(* IEC 61131-3 sources: 2026_Projet_YGO_ExcavatriceDragage/ARCHIVES/Code/MAIN, 3 files *)

(* ---- PRG_01_Inputs_LD.st ---- *)
(* ═══════════════════════════════════════════════════════════════
   📥 PRG_01_Inputs_LD — ACQUISITION & QUALIFICATION DES ENTRÉES (LADDER)
   ───────────────────────────────────────────────────────────────
   📄 Doc : DOC/AF_Partie-06_Acquisition_Qualification_IO_v2.1.md §1/§4
   ⚙️ Exécuté par la tâche PLC en position 1 (premier programme).
   🎯 Lit les 22 TOR réelles depuis leurs symboles bruts mappés (CSV
       Device_IO_20260729.csv), applique un filtre anti-rebond 20 ms et
       publie :
         • Qualified : ST_InputsQualified  (image qualifiée, lecteur unique
                                            PRG_02_Acquisition_CFC)
         • 14 scalaires legacy             (consommateurs historiques)
   🛡️ Polarité : le nom de chaque entrée dit ce que TRUE signifie. Seuls
       les freins portent InvertLogic := FALSE (REX 2026-08-03 : TRUE =
       frein OUVERT). Aucune autre inversion (contacts NC câblés 1 = sain).
   📄 Converti automatiquement en Ladder Diagram (<LD>) dans CODESYS.
   ═══════════════════════════════════════════════════════════════ *)

PROGRAM PRG_01_Inputs_LD
VAR_OUTPUT
    Qualified : ST_InputsQualified;
    PowerContactorEngaged : BOOL;   // TRUE = contacteur de puissance engagé (NO)
    EmergencyChainClosed  : BOOL;   // TRUE = boucle AU fermée (NC, câblage 1 = sain)
    PhaseRotationOk       : BOOL;   // TRUE = rotation phases correcte (NC)
    BrakeThermalFeedback  : BOOL;   // TRUE = thermique freins M1/M2/M3 OK (NC)
    M1ThermalFeedback     : BOOL;   // TRUE = thermique M1 OK (NC)
    M2ThermalFeedback     : BOOL;   // TRUE = thermique M2 OK (NC)
    M1BrakeFeedback       : BOOL;   // TRUE = frein M1 OUVERT (desserré) — REX 2026-08-03
    M2BrakeFeedback       : BOOL;   // TRUE = frein M2 OUVERT (desserré) — REX 2026-08-03
    M3BrakeFeedback       : BOOL;   // TRUE = frein M3 OUVERT (desserré) — REX 2026-08-03
    M1FwdRevSpeedFeedbackOff : BOOL; // TRUE = contacteurs sens M1 retombés (NO)
    M2FwdRevSpeedFeedbackOff : BOOL; // TRUE = contacteurs sens M2 retombés (NO)
    TopPositionSensor     : BOOL;   // TRUE = position extrême haut libre (NC)
    SlackCableSwitch      : BOOL;   // TRUE = câble M2 tendu (NC)
    KoboldContactFond     : BOOL;   // TRUE = Kobold fond détecté (NO)
END_VAR
VAR
    instPowerContactorEngaged : FB_Input;
    instEmergencyChainClosed  : FB_Input;
    instCtrlPhaseRotation     : FB_Input;
    instBrakeThermalFeedback  : FB_Input;
    instKoboldContactFond     : FB_Input;
    instHydraulicThermalOk    : FB_Input;
    instConveyorInfeedReady   : FB_Input;
    instM1FwdRevSpeedFeedbackOff : FB_Input;
    instM1Thermal             : FB_Input;
    instM1BrakeFeedback       : FB_Input;
    instM2FwdRevSpeedFeedbackOff : FB_Input;
    instM2Thermal             : FB_Input;
    instM2BrakeFeedback       : FB_Input;
    instTopPositionSensor     : FB_Input;
    instSlackCableSwitch      : FB_Input;
    instM3BrakeFeedback       : FB_Input;
    instM3ThermalFeedback     : FB_Input;
    instTranslationPosTremie  : FB_Input;
    instTranslationPosPV      : FB_Input;
    instTranslationPosP2      : FB_Input;
    instTranslationPosP1      : FB_Input;
    instTranslationPosMaintenance : FB_Input;
END_VAR

// === IMPLEMENTATION ===

// === [MACHINE] ===
// 🔌 Contacteur de puissance géré par l'arrêt d'urgence (NO) — TRUE = engagé
instPowerContactorEngaged(InputRaw := PowerContactorEngaged_DI, FilterTime := T#20MS);
PowerContactorEngaged := instPowerContactorEngaged.State;
Qualified.Machine.PowerContactorEngaged_DI := PowerContactorEngaged;

// 🔗 Boucle d'arrêt d'urgence coup-de-poing + contact PLC (NC) — TRUE = saine
instEmergencyChainClosed(InputRaw := EmergencyChainClosed_DI, FilterTime := T#20MS);
EmergencyChainClosed := instEmergencyChainClosed.State;
Qualified.Machine.EmergencyChainClosed_DI := EmergencyChainClosed;

// ⚡ Contrôle rotation phases (NC) — TRUE = correcte
instCtrlPhaseRotation(InputRaw := PhaseRotationOk_DI, FilterTime := T#20MS);
PhaseRotationOk := instCtrlPhaseRotation.State;
Qualified.Machine.PhaseRotationOk_DI := PhaseRotationOk;

// 🌡️ Thermique freins commun M1/M2/M3 (NC) — TRUE = OK
instBrakeThermalFeedback(InputRaw := BrakeThermalOk_DI, FilterTime := T#20MS);
BrakeThermalFeedback := instBrakeThermalFeedback.State;
Qualified.Machine.BrakeThermalOk_DI := BrakeThermalFeedback;

// 🪨 Détecteur fond Kobold (NO) — TRUE = fond détecté
instKoboldContactFond(InputRaw := M1_M2_KoboldContactFond_DI, FilterTime := T#20MS);
KoboldContactFond := instKoboldContactFond.State;
Qualified.Machine.M1_M2_KoboldContactFond_DI := KoboldContactFond;

// 🌡️ Thermique moteur hydraulique (NC) — TRUE = OK
instHydraulicThermalOk(InputRaw := HydraulicThermalOk_DI, FilterTime := T#20MS);
Qualified.Machine.HydraulicThermalOk_DI := instHydraulicThermalOk.State;

// ⚙️ Autorisation démarrage crible (NO) — TRUE = autorisé
instConveyorInfeedReady(InputRaw := ConveyorInfeedReady_DI, FilterTime := T#20MS);
Qualified.Machine.ConveyorInfeedReady_DI := instConveyorInfeedReady.State;

// === [WINCH] ===
// 📡 Contacteurs sens M1 relâchés (NO) — TRUE = retombés
instM1FwdRevSpeedFeedbackOff(InputRaw := M1_ContactorsReleased_DI, FilterTime := T#20MS);
M1FwdRevSpeedFeedbackOff := instM1FwdRevSpeedFeedbackOff.State;
Qualified.Winch.M1_ContactorsReleased_DI := M1FwdRevSpeedFeedbackOff;

// 🌡️ Thermique moteur M1 (NC) — TRUE = OK
instM1Thermal(InputRaw := M1_ThermalOk_DI, FilterTime := T#20MS);
M1ThermalFeedback := instM1Thermal.State;
Qualified.Winch.M1_ThermalOk_DI := M1ThermalFeedback;

// 🔒 Retour frein M1 — REX 2026-08-03 : InvertLogic := FALSE, TRUE = frein OUVERT
instM1BrakeFeedback(InputRaw := M1_BrakeIsOpen_DI, InvertLogic := FALSE, FilterTime := T#20MS);
M1BrakeFeedback := instM1BrakeFeedback.State;
Qualified.Winch.M1_BrakeIsOpen_DI := M1BrakeFeedback;

// 📡 Contacteurs sens M2 relâchés (NO) — TRUE = retombés
instM2FwdRevSpeedFeedbackOff(InputRaw := M2_ContactorsReleased_DI, FilterTime := T#20MS);
M2FwdRevSpeedFeedbackOff := instM2FwdRevSpeedFeedbackOff.State;
Qualified.Winch.M2_ContactorsReleased_DI := M2FwdRevSpeedFeedbackOff;

// 🌡️ Thermique moteur M2 (NC) — TRUE = OK
instM2Thermal(InputRaw := M2_ThermalOk_DI, FilterTime := T#20MS);
M2ThermalFeedback := instM2Thermal.State;
Qualified.Winch.M2_ThermalOk_DI := M2ThermalFeedback;

// 🔒 Retour frein M2 — REX 2026-08-03 : InvertLogic := FALSE, TRUE = frein OUVERT
instM2BrakeFeedback(InputRaw := M2_BrakeIsOpen_DI, InvertLogic := FALSE, FilterTime := T#20MS);
M2BrakeFeedback := instM2BrakeFeedback.State;
Qualified.Winch.M2_BrakeIsOpen_DI := M2BrakeFeedback;

// 🔝 Fin de course position extrême haut (NC) — TRUE = libre, déclenche AU
instTopPositionSensor(InputRaw := M1M2_TopPositionFree_DI, FilterTime := T#20MS);
TopPositionSensor := instTopPositionSensor.State;
Qualified.Winch.M1M2_TopPositionFree_DI := TopPositionSensor;

// 🔗 Capteur mou de câble M2 (NC) — TRUE = câble tendu
instSlackCableSwitch(InputRaw := M2_TensionedCable_DI, FilterTime := T#20MS);
SlackCableSwitch := instSlackCableSwitch.State;
Qualified.Winch.M2_TensionedCable_DI := SlackCableSwitch;

// === [TRANSLATION] ===
// 🔒 Retour frein M3 — REX 2026-08-03 : InvertLogic := FALSE, TRUE = frein OUVERT
instM3BrakeFeedback(InputRaw := M3_BrakeIsOpen_DI, InvertLogic := FALSE, FilterTime := T#20MS);
M3BrakeFeedback := instM3BrakeFeedback.State;
Qualified.Translation.M3_BrakeIsOpen_DI := M3BrakeFeedback;

// 🌡️ Thermique moteur M3 (NC) — TRUE = OK
instM3ThermalFeedback(InputRaw := M3_ThermalFeedback_DI, FilterTime := T#20MS);
Qualified.Translation.M3_ThermalFeedback_DI := instM3ThermalFeedback.State;

// 🏭 Capteurs de position chariot M3 (NO) — TRUE = position atteinte
instTranslationPosTremie(InputRaw := M3_PosTremie_DI, FilterTime := T#20MS);
Qualified.Translation.M3_PosTremie_DI := instTranslationPosTremie.State;

instTranslationPosPV(InputRaw := M3_PosPV_DI, FilterTime := T#20MS);
Qualified.Translation.M3_PosPV_DI := instTranslationPosPV.State;

instTranslationPosP2(InputRaw := M3_PosP2_DI, FilterTime := T#20MS);
Qualified.Translation.M3_PosP2_DI := instTranslationPosP2.State;

instTranslationPosP1(InputRaw := M3_PosP1_DI, FilterTime := T#20MS);
Qualified.Translation.M3_PosP1_DI := instTranslationPosP1.State;

instTranslationPosMaintenance(InputRaw := M3_PosMaintenance_DI, FilterTime := T#20MS);
Qualified.Translation.M3_PosMaintenance_DI := instTranslationPosMaintenance.State;

(* ---- PRG_06_Outputs_LD.st ---- *)
(* ═══════════════════════════════════════════════════════════════
   📤 PRG_06_Outputs_LD — Écriture des SORTIES physiques (PROGRAMME LADDER)
   ───────────────────────────────────────────────────────────────
   📄 Doc : DOC/AF/AF_Partie-06_Acquisition_Qualification_IO_v2.3.md §5
   ⚙️ Exécuté par la tâche PLC en position 6 (après PRG_05_Translation).
   📄 Converti automatiquement en Ladder Diagram (<LD>) dans CODESYS.
   🛡️ Barrières finales M1/M2/M3
      rendues visibles — FB_WinchOutputInterlock_LD (×2) et
      FB_TranslationOutputInterlock_LD (×1) câblés en amont des coils,
      contacts nommés sur variables qualifiées (visibilité maintenance :
      interlocks/safety qui coupent chaque actionneur lisibles directement
      dans le réseau Ladder, sans ouvrir un autre POU).
   🔒 SafetyStructureNotValidated reste TRUE : AUCUNE sortie physique
      moteur/frein n'est autorisée tant que ce garde-fou n'est pas retiré
      (voir alerte ci-dessous).
   ⚠️ FB_Safety_Winch / FB_Safety_Translation (7 mécanismes Méca A→E,
      PowerCutOff métier) ne sont pas appelés dans CODE/ : les demandes
      ST_WinchFinalInterlockRequest / ST_TranslationFinalInterlockRequest
      ne portent donc que SafeStop (partiel). Ne pas déduire que la safety
      métier complète est active.
   Coils câblées directement sur les sorties des interlocks finaux —
   simplifie la lecture maintenance.
   DriveControlWord (mot commande 0x3101) et DriveFreqRefWord (consigne
   fréquence WORD, registre 0x3100, échelle ×100 — WORD 5000 = 50,00 Hz)
   capturés en variables locales M3_DriveControlWord / M3_DriveFreqRefWord.
   Mapping E/S CODESYS (Device.export) manuel — voir §2 ci-dessous.
   ═══════════════════════════════════════════════════════════════ *)

PROGRAM PRG_06_Outputs_LD

VAR_INPUT
    // === 📥 ENTRÉES PROGRAMME (AUCUNE - REÇOIT LES ORDRES VIA PRG_04 & PRG_05) ===
END_VAR

VAR_OUTPUT
    (* Cibles de mapping : PowerKeepAliveACmd/BCmd/EmergencyArmingCmd,
       déclarées en VAR locale ci-dessous (voir §2). *)
    EmergencyArmingPulseActive   : BOOL;
    EmergencyArmingLockoutActive : BOOL;
    ArmingSeqStep                : INT;
    RedundancyTestFailed         : BOOL;
    EmergencyArmingFailed        : BOOL;
    EmergencyState               : ST_Safety_Emergency_State;
    EmergencyDiag                : ST_Safety_Emergency_Diag;
    PowerCutOffActive            : BOOL; (* TRUE = demande de coupure finale active *)

    SafetyStructureNotValidated  : BOOL := FALSE; (* 🔓 Garde-fou désactivé : les autorisations M1/M2/M3 sont liées dynamiquement à leurs sécurités *)
    // Enable ne coupe que sur PowerCutOff (barrière finale, AF02 §2, AF06 §5
    // "SafeStop laisse la décélération métier se terminer"). SafeStop est une rampe rapide
    // gérée en amont par FB_Winch/FB_Translation (Enable maintenu, AGENTS.md, TC-P03-001) ;
    // Error reflète tout ErrorId y compris les mécanismes SafeStop-only.
    M1InterlockEnable            : BOOL; (* Gate finale M1 : WinchM1FinalInterlockRequest.Enable AND NOT WinchM1FinalInterlockRequest.PowerCutOff *)
    M2InterlockEnable            : BOOL; (* Gate finale M2 : WinchM2FinalInterlockRequest.Enable AND NOT WinchM2FinalInterlockRequest.PowerCutOff *)
    M3InterlockEnable            : BOOL; (* Gate finale M3 : TranslationFinalInterlockRequest.Enable AND NOT TranslationFinalInterlockRequest.PowerCutOff *)
    // Réseau informatif séparé : visibilité maintenance de ce qui
    // bloque (PowerCutOff / SafeStop / Global), SANS influencer Enable — juste de l'information en Watch/Ladder.
    M1PowerCutOffSafetyInfo      : BOOL;
    M1SafeStopSafetyInfo         : BOOL;
    M1BlockedBySafetyInfo        : BOOL;

    M2PowerCutOffSafetyInfo      : BOOL;
    M2SafeStopSafetyInfo         : BOOL;
    M2BlockedBySafetyInfo        : BOOL;

    M3PowerCutOffSafetyInfo      : BOOL;
    M3SafeStopSafetyInfo         : BOOL;
    M3BlockedBySafetyInfo        : BOOL;

    (* Les noms Device bruts ( *_DQ / *_RQ ), ex. M1_RelayFwd_Up_DQ,
       M3_BrakeRelease_RQ) ne sont pas déclarés ici : les déclarer créerait une collision
       de portée avec la variable GLOBALE homonyme créée par le mapping E/S CODESYS
       (Device.export), qui masquerait le pilotage matériel réel (voir §2 plus bas
       pour le détail et la liste des chemins qualifiés à mapper). *)
    TranslationBrakeCmd          : BOOL; // <-- [ACT] Demande frein M3 arbitree — cible du mapping E/S
    M3_DriveControlWord          : WORD; // <-- [ACT] Mot de commande variateur M3 (0x3101) — cible du mapping E/S
    M3_DriveFreqRefWord          : WORD; // <-- [ACT] Consigne frequence variateur M3 (0x3100, x100) — cible du mapping E/S

    // === ⚡ ORDRES ACTIONNEURS (ACCESSIBLES SIMULATION / PROCESS) ===
    M1RelayFwd                   : BOOL; // <-- [ACT] Ordre contacteur montee treuil M1
    M1RelayRev                   : BOOL; // <-- [ACT] Ordre contacteur descente treuil M1
    M1SpeedContactor1            : BOOL; // <-- [ACT] Ordre contacteur palier 1 treuil M1
    M1SpeedContactor2            : BOOL; // <-- [ACT] Ordre contacteur palier 2 treuil M1
    M1SpeedContactor3            : BOOL; // <-- [ACT] Ordre contacteur palier 3 treuil M1
    M1SpeedContactor4            : BOOL; // <-- [ACT] Ordre contacteur palier 4 treuil M1
    M1BrakeCmd                   : BOOL; // <-- [ACT] Ordre desserrage frein M1 (1=Desserrer)
    M2RelayFwd                   : BOOL; // <-- [ACT] Ordre contacteur montee/fermeture treuil M2
    M2RelayRev                   : BOOL; // <-- [ACT] Ordre contacteur descente/ouverture treuil M2
    M2SpeedContactor1            : BOOL; // <-- [ACT] Ordre contacteur palier 1 treuil M2
    M2SpeedContactor2            : BOOL; // <-- [ACT] Ordre contacteur palier 2 treuil M2
    M2SpeedContactor3            : BOOL; // <-- [ACT] Ordre contacteur palier 3 treuil M2
    M2SpeedContactor4            : BOOL; // <-- [ACT] Ordre contacteur palier 4 treuil M2
    M2BrakeCmd                   : BOOL; // <-- [ACT] Ordre desserrage frein M2 (1=Desserrer)
    KoboldContactorCmd           : BOOL; // <-- [ACT] Ordre alimentation contacteur capteur fond Kobold
    PowerKeepAliveACmd           : BOOL; // <-- [SAFE] Maintien puissance voie A (1=Maintenu)
    PowerKeepAliveBCmd           : BOOL; // <-- [SAFE] Maintien puissance voie B (1=Maintenu)
    EmergencyArmingCmd           : BOOL; // <-- [CMD] Impulsion rearmement puissance AU
END_VAR

VAR
    // === 🛡️ SOUS-INSTANCES FB INTERLOCKS SORTIES ===
    instWinchOutputInterlockM1       : FB_WinchOutputInterlock_LD;       // * [INST] Barriere finale treuil M1
    instWinchOutputInterlockM2       : FB_WinchOutputInterlock_LD;       // * [INST] Barriere finale treuil M2
    instTranslationOutputInterlockM3 : FB_TranslationOutputInterlock_LD; // * [INST] Barriere finale translation M3
    instSafetyEmergencyManagement    : FB_Safety_EmergencyManagement;    // * [INST] Gestionnaire de rearmement AU

    // === ⚙️ VARIABLES LOCALES INTERNES ===
    PowerCutOffReq                   : BOOL; // . [LOC] Demande agregative coupure puissance
END_VAR

// === 🛡️ §1 BARRIÈRES FINALES M1 / M2 / M3 — INTERLOCKS VISIBLES ===
// Chaque bloc reçoit la demande brute publique du procédé propriétaire
// (ST_WinchFinalInterlockRequest / ST_TranslationFinalInterlockRequest) :
// tous les interlocks/safety qui peuvent couper cet actionneur sont donc
// lisibles directement sur ce réseau, sans ouvrir un autre POU.

// ── Interlock final M1 (Treuil Retenue) ──────────────────────────────────
M1InterlockEnable := PRG_04_Treuils_Benne.WinchM1FinalInterlockRequest.Enable
                      AND NOT PRG_04_Treuils_Benne.WinchM1FinalInterlockRequest.PowerCutOff;

// Info diagnostic seule (Watch/Ladder) — ne participe PAS au calcul ci-dessus.
// 🧨 Bloc 1 : Sécurités entraînant un PowerCutOff (coupure puissance)
M1PowerCutOffSafetyInfo := OR(
    PRG_04_Treuils_Benne.WinchM1Safety.PowerCutOff,
    PRG_04_Treuils_Benne.WinchM1Safety.ErrorMecaA,
    PRG_04_Treuils_Benne.WinchM1Safety.ErrorMecaB,
    PRG_04_Treuils_Benne.WinchM1Safety.ErrorMecaC,
    PRG_04_Treuils_Benne.WinchM1Safety.ErrorMecaD,
    PRG_04_Treuils_Benne.WinchM1Safety.ErrorMecaE,
    PRG_04_Treuils_Benne.WinchM1Safety.ThermalFault
);

// 🛡️ Bloc 2 : Défauts sécurité entraînant un SafeStop / Rampe rapide
M1SafeStopSafetyInfo := OR(
    PRG_04_Treuils_Benne.WinchM1Safety.SafeStop,
    PRG_04_Treuils_Benne.WinchM1Safety.Error,
    PRG_04_Treuils_Benne.WinchM1Safety.ErrorOperatorComm,
    PRG_04_Treuils_Benne.WinchM1Safety.ErrorEncoder,
    PRG_04_Treuils_Benne.WinchM1Safety.ErrorPhaseRotation,
    PRG_04_Treuils_Benne.WinchM1Safety.ErrorOppositeDir,
    PRG_04_Treuils_Benne.WinchM1Safety.ErrorNoMovement
);

// 🚫 Bloc 3 : Synthèse globale du blocage sécurité (PowerCutOff OU SafeStop)
M1BlockedBySafetyInfo := OR(
    M1PowerCutOffSafetyInfo,
    M1SafeStopSafetyInfo
);

instWinchOutputInterlockM1(
    Enable                     := M1InterlockEnable,
    Reset                      := PRG_07_Supervision.FaultMachineReset_IHM,
    PowerContactorEngaged      := PRG_04_Treuils_Benne.WinchM1FinalInterlockRequest.PowerContactorEngaged,
    SafeStop                   := PRG_04_Treuils_Benne.WinchM1FinalInterlockRequest.SafeStop,
    BrakeFeedback              := PRG_04_Treuils_Benne.WinchM1FinalInterlockRequest.BrakeFeedback,
    FwdRevSpeedFeedbackOff     := PRG_04_Treuils_Benne.WinchM1FinalInterlockRequest.FwdRevSpeedFeedbackOff,
    RequestedRelayFwd          := PRG_04_Treuils_Benne.WinchM1FinalInterlockRequest.RequestedRelayFwd,
    RequestedRelayRev          := PRG_04_Treuils_Benne.WinchM1FinalInterlockRequest.RequestedRelayRev,
    RequestedContactor1        := PRG_04_Treuils_Benne.WinchM1FinalInterlockRequest.RequestedContactor1,
    RequestedContactor2        := PRG_04_Treuils_Benne.WinchM1FinalInterlockRequest.RequestedContactor2,
    RequestedContactor3        := PRG_04_Treuils_Benne.WinchM1FinalInterlockRequest.RequestedContactor3,
    RequestedContactor4        := PRG_04_Treuils_Benne.WinchM1FinalInterlockRequest.RequestedContactor4,
    RequestedStep               := PRG_04_Treuils_Benne.WinchM1FinalInterlockRequest.RequestedStep
);

M1RelayFwd        := instWinchOutputInterlockM1.RelayFwd;
M1RelayRev        := instWinchOutputInterlockM1.RelayRev;
M1SpeedContactor1 := instWinchOutputInterlockM1.Contactor1;
M1SpeedContactor2 := instWinchOutputInterlockM1.Contactor2;
M1SpeedContactor3 := instWinchOutputInterlockM1.Contactor3;
M1SpeedContactor4 := instWinchOutputInterlockM1.Contactor4;
// Recalcul INDEPENDANT sur les DQ
// finaux (pas une simple recopie de instWinchOutputInterlockM1.BrakeCmd) -- visible ici
// sans ouvrir FB_WinchOutputInterlock_LD, meme doctrine que le reste de ce POU.
M1BrakeCmd        := M1RelayFwd OR M1RelayRev;

// ── Interlock final M2 (Treuil Benne) ────────────────────────────────────
M2InterlockEnable := PRG_04_Treuils_Benne.WinchM2FinalInterlockRequest.Enable
                      AND NOT PRG_04_Treuils_Benne.WinchM2FinalInterlockRequest.PowerCutOff;

// Info diagnostic seule (Watch/Ladder) — ne participe PAS au calcul ci-dessus.
// 🧨 Bloc 1 : Sécurités entraînant un PowerCutOff (coupure puissance)
M2PowerCutOffSafetyInfo := OR(
    PRG_04_Treuils_Benne.WinchM2Safety.PowerCutOff,
    PRG_04_Treuils_Benne.WinchM2Safety.ErrorMecaA,
    PRG_04_Treuils_Benne.WinchM2Safety.ErrorMecaB,
    PRG_04_Treuils_Benne.WinchM2Safety.ErrorMecaC,
    PRG_04_Treuils_Benne.WinchM2Safety.ErrorMecaD,
    PRG_04_Treuils_Benne.WinchM2Safety.ErrorMecaE,
    PRG_04_Treuils_Benne.WinchM2Safety.ThermalFault
);

// 🛡️ Bloc 2 : Défauts sécurité entraînant un SafeStop / Rampe rapide / Verrous Benne
M2SafeStopSafetyInfo := OR(
    PRG_04_Treuils_Benne.WinchM2Safety.SafeStop,
    PRG_04_Treuils_Benne.WinchM2Safety.Error,
    PRG_04_Treuils_Benne.WinchM2Safety.ErrorOperatorComm,
    PRG_04_Treuils_Benne.WinchM2Safety.ErrorEncoder,
    PRG_04_Treuils_Benne.WinchM2Safety.ErrorPhaseRotation,
    PRG_04_Treuils_Benne.WinchM2Safety.ErrorOppositeDir,
    PRG_04_Treuils_Benne.WinchM2Safety.ErrorNoMovement,
    PRG_04_Treuils_Benne.WinchM2Safety.SlackCable,
    PRG_04_Treuils_Benne.BucketState.Error,
    PRG_04_Treuils_Benne.BucketState.CoupledMotionBlockedByBucket
);

// 🚫 Bloc 3 : Synthèse globale du blocage sécurité (PowerCutOff OU SafeStop)
M2BlockedBySafetyInfo := OR(
    M2PowerCutOffSafetyInfo,
    M2SafeStopSafetyInfo
);

instWinchOutputInterlockM2(
    Enable                     := M2InterlockEnable,
    Reset                      := PRG_07_Supervision.FaultMachineReset_IHM,
    PowerContactorEngaged      := PRG_04_Treuils_Benne.WinchM2FinalInterlockRequest.PowerContactorEngaged,
    SafeStop                   := PRG_04_Treuils_Benne.WinchM2FinalInterlockRequest.SafeStop,
    BrakeFeedback              := PRG_04_Treuils_Benne.WinchM2FinalInterlockRequest.BrakeFeedback,
    FwdRevSpeedFeedbackOff     := PRG_04_Treuils_Benne.WinchM2FinalInterlockRequest.FwdRevSpeedFeedbackOff,
    RequestedRelayFwd          := PRG_04_Treuils_Benne.WinchM2FinalInterlockRequest.RequestedRelayFwd,
    RequestedRelayRev          := PRG_04_Treuils_Benne.WinchM2FinalInterlockRequest.RequestedRelayRev,
    RequestedContactor1        := PRG_04_Treuils_Benne.WinchM2FinalInterlockRequest.RequestedContactor1,
    RequestedContactor2        := PRG_04_Treuils_Benne.WinchM2FinalInterlockRequest.RequestedContactor2,
    RequestedContactor3        := PRG_04_Treuils_Benne.WinchM2FinalInterlockRequest.RequestedContactor3,
    RequestedContactor4        := PRG_04_Treuils_Benne.WinchM2FinalInterlockRequest.RequestedContactor4,
    RequestedStep               := PRG_04_Treuils_Benne.WinchM2FinalInterlockRequest.RequestedStep
);

M2RelayFwd        := instWinchOutputInterlockM2.RelayFwd;
M2RelayRev        := instWinchOutputInterlockM2.RelayRev;
M2SpeedContactor1 := instWinchOutputInterlockM2.Contactor1;
M2SpeedContactor2 := instWinchOutputInterlockM2.Contactor2;
M2SpeedContactor3 := instWinchOutputInterlockM2.Contactor3;
M2SpeedContactor4 := instWinchOutputInterlockM2.Contactor4;
// Recalcul INDEPENDANT, voir M1 ci-dessus.
M2BrakeCmd        := M2RelayFwd OR M2RelayRev;

// KoboldContactorCmd est écrit depuis la commande arbitrée
// PRG_04_Treuils_Benne.KoboldContactorCmdArbitrated. Mapping E/S CODESYS
// (voir §2 plus bas) : M1_M2_KoboldMeasureEnable_DQ <- PRG_06_Outputs_LD.KoboldContactorCmd.
KoboldContactorCmd := PRG_04_Treuils_Benne.KoboldContactorCmdArbitrated;

// ── Interlock final M3 (Translation, variateur AC600) ────────────────────
// 🛡️ Déblocage M3 sans forçage manuel de SafetyStructureNotValidated.
// Ne coupe que sur PowerCutOff — voir commentaire VAR_OUTPUT en tête de fichier.
M3InterlockEnable := PRG_05_Translation.TranslationFinalInterlockRequest.Enable
                      AND NOT PRG_05_Translation.TranslationFinalInterlockRequest.PowerCutOff;

// Info diagnostic seule (Watch/Ladder) — ne participe PAS au calcul ci-dessus.
// 🧨 Bloc 1 : Sécurités entraînant un PowerCutOff (coupure puissance)
M3PowerCutOffSafetyInfo := OR(
    PRG_05_Translation.TranslationSafety.PowerCutOff,
    PRG_05_Translation.TranslationSafety.ErrorMecaA,
    PRG_05_Translation.TranslationSafety.ErrorMecaB,
    PRG_05_Translation.TranslationSafety.ErrorBrakeThermal
);

// 🛡️ Bloc 2 : Défauts sécurité entraînant un SafeStop / Rampe rapide
M3SafeStopSafetyInfo := OR(
    PRG_05_Translation.TranslationSafety.SafeStop,
    PRG_05_Translation.TranslationSafety.Error,
    PRG_05_Translation.TranslationSafety.ErrorOperatorComm,
    PRG_05_Translation.TranslationSafety.ErrorDriveComm,
    PRG_05_Translation.TranslationSafety.ErrorPhaseRotation,
    PRG_05_Translation.TranslationSafety.ErrorLimitSwitch,
    PRG_05_Translation.TranslationSafety.ErrorSensorIncoherent
);

// 🚫 Bloc 3 : Synthèse globale du blocage sécurité (PowerCutOff OU SafeStop)
M3BlockedBySafetyInfo := OR(
    M3PowerCutOffSafetyInfo,
    M3SafeStopSafetyInfo
);

instTranslationOutputInterlockM3(
    Enable                     := M3InterlockEnable,
    Reset                      := PRG_07_Supervision.FaultMachineReset_IHM,
    PowerContactorEngaged      := PRG_05_Translation.TranslationFinalInterlockRequest.PowerContactorEngaged,
    SafeStop                   := PRG_05_Translation.TranslationFinalInterlockRequest.SafeStop,
    BrakeReleaseRequest        := PRG_05_Translation.TranslationFinalInterlockRequest.BrakeReleaseRequest,
    BrakeCommandOpenConfirmed  := PRG_05_Translation.TranslationFinalInterlockRequest.BrakeCommandOpenConfirmed,
    RequestedDriveControlWord  := PRG_05_Translation.TranslationFinalInterlockRequest.RequestedDriveControlWord,
    RequestedDriveFreqHz       := PRG_05_Translation.TranslationFinalInterlockRequest.RequestedDriveFreqHz
);

TranslationBrakeCmd := instTranslationOutputInterlockM3.BrakeCmd;
M3_CommandWord := instTranslationOutputInterlockM3.DriveControlWord;
M3_SetpointFrequencyHz := instTranslationOutputInterlockM3.DriveFreqRefWord;

// === ⚡ §2 SORTIES PHYSIQUES DIRECTES (M1 / M2 / M3 / AU / KOBOLD) — COILS HW ===
// Pilotage direct des variables de mapping E/S matérielles :
M1_RelayFwd_Up_DQ            := M1RelayFwd;
M1_RelayRev_Down_DQ          := M1RelayRev;
M1_SpeedContactor_1_DQ       := M1SpeedContactor1;
M1_SpeedContactor_2_DQ       := M1SpeedContactor2;
M1_SpeedContactor_3_DQ       := M1SpeedContactor3;
M1_SpeedContactor_4_DQ       := M1SpeedContactor4;
M1_BrakeRelease_RQ           := M1BrakeCmd;

M2_RelayFwd_Up_Close_DQ      := M2RelayFwd;
M2_RelayRev_Down_Open_DQ     := M2RelayRev;
M2_SpeedContactor_1_DQ       := M2SpeedContactor1;
M2_SpeedContactor_2_DQ       := M2SpeedContactor2;
M2_SpeedContactor_3_DQ       := M2SpeedContactor3;
M2_SpeedContactor_4_DQ       := M2SpeedContactor4;
M2_BrakeRelease_RQ           := M2BrakeCmd;

M3_BrakeRelease_RQ           := TranslationBrakeCmd;

M1_M2_KoboldMeasureEnable_DQ := KoboldContactorCmd;

PowerKeepAlive_A_RQ          := PowerKeepAliveACmd;
PowerKeepAlive_B_RQ          := PowerKeepAliveBCmd;
EmergencyArming_RQ           := EmergencyArmingCmd;

// === 🛡️ §3 SÉCURITÉ & COUPURE PUISSANCE AMONT ===

// PowerCutOffReq = agrégation OU strict des demandes de coupure des trois procédés (M5, A-04) :
//   PowerCutOffReq = WinchM1FinalInterlockRequest.PowerCutOff
//                  OR WinchM2FinalInterlockRequest.PowerCutOff
//                  OR TranslationFinalInterlockRequest.PowerCutOff
// ⚠️ Cette ligne ST est UNIQUEMENT documentaire (contrat fonctionnel) : PRG_06_Outputs_LD est
// intégralement généré par l'oracle Python (gen_prg06_oracle.py). Contrat réel, câblé dans
// l'oracle (3 contacts parallèles sur la même coil PowerCutOffReq, voir section PowerCutOffReq
// du script).
PowerCutOffReq := PRG_05_Translation.TranslationFinalInterlockRequest.PowerCutOff;

instSafetyEmergencyManagement(
    Enable := TRUE,
    Reset := PRG_07_Supervision.FaultMachineReset_IHM,
    ArmRequest := GVL_IHM.Modes.Cmd.BtnEmergencyArming,
    EmergencyChainClosed := PRG_02_Acquisition.HwIn.Machine.EmergencyChainClosed_DI,
    PowerContactorEngaged := PRG_02_Acquisition.HwIn.Machine.PowerContactorEngaged_DI,
    PowerCutOffRequest := PowerCutOffReq,
    BtnEmergencyCutOff := GVL_IHM.Modes.Cmd.BtnEmergencyCutOff
);

PowerKeepAliveACmd := instSafetyEmergencyManagement.MaintainA_RQ;
PowerKeepAliveBCmd := instSafetyEmergencyManagement.MaintainB_RQ;
EmergencyArmingCmd := instSafetyEmergencyManagement.ArmPulse_RQ;

EmergencyArmingLockoutActive := instSafetyEmergencyManagement.EmergencyArmingLockoutActive;
ArmingSeqStep := instSafetyEmergencyManagement.ArmingSeqStep;
RedundancyTestFailed := instSafetyEmergencyManagement.RedundancyTestFailed;
EmergencyArmingFailed := instSafetyEmergencyManagement.EmergencyArmingFailed;
EmergencyState := instSafetyEmergencyManagement.State;
EmergencyDiag := instSafetyEmergencyManagement.Diag;
PowerCutOffActive := PowerCutOffReq;

END_PROGRAM

(* ---- PRG_ACQUISITION_CFC.st ---- *)
(* ═══════════════════════════════════════════════════════════════
   📡 PRG_ACQUISITION_CFC — Acquisition brute, simulation et aiguillage HwIn
   ───────────────────────────────────────────────────────────────
   📄 Docs : DOC/AF_Partie-06_Acquisition_Qualification_IO_v2.0.md §2 ;
            DOC/AF_Partie-13_Fonction_Simulation_v2.0.md
   ⚙️ Version ST temporaire pour validation (cible CFC).
   🎯 Rôle unique : produire l'image matérielle HwIn consommée par le reste
      du programme. Aucune décision métier (SafeStop, mode, commande) ici.
   🔗 Producteur unique de HwIn ; consommateurs = PRG_INPUTS_LD et suivants.
   ═══════════════════════════════════════════════════════════════ *)

PROGRAM PRG_ACQUISITION_CFC

VAR_OUTPUT
    HwReal                   : ST_HardwareImage;  (* Image matérielle brute lue sur le terrain *)
    HwSim                    : ST_HardwareImage;  (* Image produite par le banc de simulation *)
    HwIn                     : ST_HardwareImage;  (* Image aiguillée réel/simulé *)
    WinchInputSourceChanged  : BOOL;              (* Pulse 1 cycle sur bascule réel/simulé domaine Winch *)

    // 🆕 Migration PRG_00_Inputs : positions Translation M3 exposées en sortie de programme
    TranslationPosTremie      : BOOL;   (* TRUE = translation en position Trémie *)
    TranslationPosPV          : BOOL;   (* TRUE = translation en zone pré-ralentissement PV *)
    TranslationPosP2          : BOOL;   (* TRUE = translation en position P2 *)
    TranslationPosP1          : BOOL;   (* TRUE = translation en position P1 *)
    TranslationPosMaintenance : BOOL;   (* TRUE = translation en position Maintenance *)

    // 🆕 Migration PRG_00_Inputs : retours variateur M3 filtrés (PT1 T#0MS = recopie legacy)
    M3_StatusWord_Filtered        : UINT;
    M3_ActualFrequencyHz_Filtered : UINT;
END_VAR

VAR
    (* ── Instances de traitement complexes ── *)
    instSimBench             : FB_SimBench;
    instJoystick             : FB_Joystick;
    instEncoderAbsM1         : FB_Encoder_Abs;
    instEncoderScaleM1       : FB_Encoder_Scale;
    instHomingM1             : FB_Encoder_Homing;
    instEncoderAbsM2         : FB_Encoder_Abs;
    instEncoderScaleM2       : FB_Encoder_Scale;
    instHomingM2             : FB_Encoder_Homing;
    instPosDecoderM3         : FB_Translation_PositionDecoder;

    (* ── Filtrage des retours variateur M3 (migration PRG_00_Inputs) ── *)
    instCycleTimeAcq            : FB_CycleTime;
    instFilterM3StatusWord      : FB_Filter_PT1;
    instFilterM3ActualFreqHz      : FB_Filter_PT1;

    (* ── Mémoire de la source Winch (front bascule réel/simulé) ── *)
    WinchInputSourceSimulated            : BOOL;
    PreviousWinchInputSourceSimulated    : BOOL;
    WinchInputSourceInitialized          : BOOL;
END_VAR

// === IMPLEMENTATION ===

// ─── §0 MATÉRIEL ──► HwReal (Acquisition brute unique) ─────────────────────────

// Winch M1 / M2 et codeurs
HwReal.Winch.M1_ContactorsReleased_DI := M1_ContactorsReleased_DI;
HwReal.Winch.M1_ThermalOk_DI          := M1_ThermalOk_DI;
HwReal.Winch.M1_BrakeIsOpen_DI        := M1_BrakeIsOpen_DI;

HwReal.Winch.M2_ContactorsReleased_DI := M2_ContactorsReleased_DI;
HwReal.Winch.M2_ThermalOk_DI          := M2_ThermalOk_DI;
HwReal.Winch.M2_BrakeIsOpen_DI        := M2_BrakeIsOpen_DI;

HwReal.Winch.M1M2_TopPositionFree_DI  := M1M2_TopPositionFree_DI;
HwReal.Winch.M2_TensionedCable_DI     := M2_TensionedCable_DI;

HwReal.Winch.COD1_PosValue            := COD1_PosValue;
HwReal.Winch.COD1_Alarms              := COD1_Alarms;
HwReal.Winch.COD1_Warnings            := COD1_Warnings;
HwReal.Winch.COD1_DeviceState         := COD1_CODEUR.GetDeviceState();

HwReal.Winch.COD2_PosValue            := COD2_PosValue;
HwReal.Winch.COD2_Alarms              := COD2_Alarms;
HwReal.Winch.COD2_Warnings            := COD2_Warnings;
HwReal.Winch.COD2_DeviceState         := COD2_CODEUR.GetDeviceState();

// Translation M3 et variateur AC600
HwReal.Translation.M3_PosTremie_DI      := M3_PosTremie_DI;
HwReal.Translation.M3_PosPV_DI          := M3_PosPV_DI;
HwReal.Translation.M3_PosP2_DI          := M3_PosP2_DI;
HwReal.Translation.M3_PosP1_DI          := M3_PosP1_DI;
HwReal.Translation.M3_PosMaintenance_DI := M3_PosMaintenance_DI;
HwReal.Translation.M3_BrakeIsOpen_DI    := M3_BrakeIsOpen_DI;
HwReal.Translation.M3_ThermalFeedback_DI:= M3_ThermalFeedback_DI; // 🆕 T96 — diagnostic seul (voie déjà mappée CODESYS, jamais lue jusqu'ici)
HwReal.Translation.M3_StatusWord        := M3_StatusWord;
HwReal.Translation.M3_ActualFrequencyHz := M3_ActualFrequencyHz;
HwReal.Translation.AC600_DeviceState    := AC600_ECAT_Drive.GetDeviceState();

// Opérateur / Joystick / bus CANopen
HwReal.Operator.JoyXRaw_ANA1      := JoyXRaw_ANA1;
HwReal.Operator.JoyYRaw_ANA2      := JoyYRaw_ANA2;
HwReal.Operator.JoyBtnRaw         := JoyBtnRaw;
HwReal.Operator.CanBusState       := CANbus.GetBusState();
HwReal.Operator.JOY1_DeviceState  := JOY1_JOYSTICK_MCB560_CO4201A.GetDeviceState();

// Sécurités / Communs Machine
HwReal.Machine.PowerContactorEngaged_DI   := PowerContactorEngaged_DI;
HwReal.Machine.EmergencyChainClosed_DI    := EmergencyChainClosed_DI;
HwReal.Machine.PhaseRotationOk_DI         := PhaseRotationOk_DI;
HwReal.Machine.BrakeThermalOk_DI          := BrakeThermalOk_DI;
HwReal.Machine.M1_M2_KoboldContactFond_DI := M1_M2_KoboldContactFond_DI;
HwReal.Machine.HydraulicThermalOk_DI      := HydraulicThermalOk_DI;

// ─── §0bis HwReal / SimBench ──► HwIn (Aiguillage simulation par domaine) ──────

instSimBench(
    Enable                   := GVL_Simulation.SimulationModeActive,
    M1_RelayFwd              := GVL_Global.M1RelayFwd,
    M1_RelayRev              := GVL_Global.M1RelayRev,
    M1_SpeedContactor_1      := GVL_Global.M1SpeedContactor1,
    M1_SpeedContactor_2      := GVL_Global.M1SpeedContactor2,
    M1_SpeedContactor_3      := GVL_Global.M1SpeedContactor3,
    M1_SpeedContactor_4      := GVL_Global.M1SpeedContactor4,
    M1_SpeedRefPct           := PRG_TREUILS_CFC.M1_SpeedRef_Active,
    M1_PresetTriggerCmd      := PRG_02_Encoders.instEncoderAbsM1.PresetTriggerCmd,
    M1_PresetValueOut        := PRG_02_Encoders.instEncoderAbsM1.PresetValueOut,
    M1_BrakeCmd              := GVL_Global.M1BrakeCmd,
    M2_RelayFwd              := GVL_Global.M2RelayFwd,
    M2_RelayRev              := GVL_Global.M2RelayRev,
    M2_SpeedContactor_1      := GVL_Global.M2SpeedContactor1,
    M2_SpeedContactor_2      := GVL_Global.M2SpeedContactor2,
    M2_SpeedContactor_3      := GVL_Global.M2SpeedContactor3,
    M2_SpeedContactor_4      := GVL_Global.M2SpeedContactor4,
    M2_SpeedRefPct           := PRG_TREUILS_CFC.M2_SpeedRef_Active,
    M2_PresetTriggerCmd      := PRG_02_Encoders.instEncoderAbsM2.PresetTriggerCmd,
    M2_PresetValueOut        := PRG_02_Encoders.instEncoderAbsM2.PresetValueOut,
    M2_BrakeCmd              := GVL_Global.M2BrakeCmd,
    M3_Direction             := PRG_TRANSLATION_CFC.M3_Direction_Active,
    M3_SpeedRefPct           := PRG_TRANSLATION_CFC.M3_SpeedRef_Active,
    M3_BrakeCmd              := GVL_Global.TranslationBrakeCmd,
    M3_TargetNum             := GVL_IHM.TranslationM3.Cmd.SelTarget,
    PowerKeepAlive_A         := PRG_10_Outputs_LD.PowerKeepAlive_A_RQ,
    PowerKeepAlive_B         := PRG_10_Outputs_LD.PowerKeepAlive_B_RQ,
    EmergencyArming_RQ       := PRG_10_Outputs_LD.EmergencyArming_RQ,
    SimEncoderSpeedFactor    := GVL_Simulation.SimEncoderSpeedFactor,
    SimSyncDeviationInjectM1 := GVL_Simulation.SimSyncDeviationInjectM1,
    SimSyncDeviationInjectM2 := GVL_Simulation.SimSyncDeviationInjectM2,
    SimSyncDeviationOffset_M := GVL_Simulation.SimSyncDeviationOffset_M,
    SimM3SensorsWordActive   := GVL_Simulation.SimM3SensorsWordActive,
    SimM3SensorsWord         := GVL_Simulation.SimM3SensorsWord,
    SimJoystickRawX          := GVL_Simulation.SimJoystickRawX,
    SimJoystickRawY          := GVL_Simulation.SimJoystickRawY,
    SimJoystickRawButton     := GVL_Simulation.SimJoystickRawButton,
    SimKoboldContactValue    := GVL_Simulation.SimKoboldContactValue,
    BtnEmergencyStop         := GVL_IHM.Modes.Cmd.BtnEmergencyCutOff,
    HwReal                   := HwReal,
    RawPosM1                 := _SimEncoderRawPosM1,
    RawPosM2                 := _SimEncoderRawPosM2
);

// 🧪 Image du banc exposée pour lecture côte à côte ; aucune logique métier ne lit HwSim.
HwSim.Winch       := instSimBench.Winch;
HwSim.Translation := instSimBench.Translation;
HwSim.Operator    := instSimBench.Operator;
HwSim.Machine     := instSimBench.Machine;

// 🔄 Source Winch atomique + pulse générique. Au boot, la source initiale est mémorisée sans faux pulse.
WinchInputSourceSimulated := GVL_Simulation.SimulationModeActive AND GVL_Simulation.SimWinchActive;
IF NOT WinchInputSourceInitialized THEN
    PreviousWinchInputSourceSimulated := WinchInputSourceSimulated;
    WinchInputSourceInitialized := TRUE;
    WinchInputSourceChanged := FALSE;
ELSE
    WinchInputSourceChanged := (WinchInputSourceSimulated <> PreviousWinchInputSourceSimulated);
    PreviousWinchInputSourceSimulated := WinchInputSourceSimulated;
END_IF;

// Aiguillage domaine par domaine (réel si simulateur inactif pour ce domaine).
IF WinchInputSourceSimulated
    THEN HwIn.Winch := instSimBench.Winch;             ELSE HwIn.Winch := HwReal.Winch;             END_IF;
IF GVL_Simulation.SimulationModeActive AND GVL_Simulation.SimTranslationActive
    THEN HwIn.Translation := instSimBench.Translation; ELSE HwIn.Translation := HwReal.Translation; END_IF;
IF GVL_Simulation.SimulationModeActive AND GVL_Simulation.SimOperatorActive
    THEN HwIn.Operator := instSimBench.Operator;       ELSE HwIn.Operator := HwReal.Operator;       END_IF;
IF GVL_Simulation.SimulationModeActive AND GVL_Simulation.SimMachineActive
    THEN HwIn.Machine := instSimBench.Machine;         ELSE HwIn.Machine := HwReal.Machine;         END_IF;

// ─── §1 TRAITEMENT DES ENTRÉES COMPLEXES (depuis HwIn) ───────────────────────

// 🕹️ Joystick : acquisition + homme-mort + mise à l'échelle
instJoystick(
    Enable                    := TRUE,
    Reset                     := PRG_SUPERVISION_CFC.FaultMachineReset_IHM,
    PowerContactorEngaged     := HwIn.Machine.PowerContactorEngaged_DI,
    Mode                      := PRG_MODES_CFC.Auth.Mode,
    BenneBusy                 := PRG_TREUILS_CFC.instBucket.Busy,
    PreserveArmingAfterBucket := PRG_TREUILS_CFC.instExtractionSequence.Busy
                                 AND (PRG_TREUILS_CFC.instExtractionSequence.ExtractionState = E_ExtractionSequenceState.CLOSING_BUCKET),
    BusCanOpenOP              := PRG_01_Diagnostics.instDiagCanOpen.DeviceCanOpenMaster,
    JoystickOP                := PRG_01_Diagnostics.instDiagCanOpen.DeviceJoystick,
    RawX                      := HwIn.Operator.JoyXRaw_ANA1,
    RawY                      := HwIn.Operator.JoyYRaw_ANA2,
    RawButton                 := HwIn.Operator.JoyBtnRaw,
    BtnCalibrate              := GVL_IHM.JOY1Joystick.Cmd.BtnCalibrate,
    InvertX                   := _JoystickInvertX,
    InvertY                   := _JoystickInvertY,
    Deadband                  := _JoystickDeadband_Pct,
    FilterTime                := _JoystickFilterTime,
    DeadmanRearmTimeout       := T#10S,
    NeutralHoldTime           := T#500MS,
    NeutralXMem               := _JoystickNeutralX,
    NeutralYMem               := _JoystickNeutralY
);

// 🧲 Codeurs M1 : Abs → Homing → Scale
instEncoderAbsM1(
    Enable              := TRUE,
    Reset               := PRG_SUPERVISION_CFC.FaultMachineReset_IHM,
    PowerContactorEngaged     := HwIn.Machine.PowerContactorEngaged_DI,
    Mode                := PRG_MODES_CFC.Auth.Mode,
    RawPosIn            := HwIn.Winch.COD1_PosValue,
    AlarmsIn            := HwIn.Winch.COD1_Alarms,
    WarningsIn          := HwIn.Winch.COD1_Warnings,
    SlaveOperational    := PRG_01_Diagnostics.instDiagEthercat.DeviceEncoderM1.Operational,
    PresetRequest       := instHomingM1.PresetRequest,
    PresetValue         := instHomingM1.PresetValue
);

instHomingM1(
    Enable               := TRUE,
    Reset                := PRG_SUPERVISION_CFC.FaultMachineReset_IHM,
    PowerContactorEngaged      := HwIn.Machine.PowerContactorEngaged_DI,
    Mode                 := PRG_MODES_CFC.Auth.Mode,
    Home                 := GVL_IHM.M1TreuilRetenue.Cmd.BtnHome OR GVL_IHM.M1TreuilRetenue.Cmd.BtnHomingAtZero,
    UnitaryMode          := (PRG_MODES_CFC.Auth.Mode = E_Mode.MAINT_N2)
                            AND (PRG_MODES_CFC.Auth.JoystickWinchSelectArbitrated <> 3),
    WinchSelected        := (PRG_MODES_CFC.Auth.JoystickWinchSelectArbitrated = 1),
    CfgHomingTargetM        := _WinchM1CfgPersist.CfgHomingTarget_M,
    BtnConfirmCoherence     := GVL_IHM.M1TreuilRetenue.Cmd.BtnConfirmCoherence,
    TopPositionSensor    := HwIn.Winch.M1M2_TopPositionFree_DI,
    CfgTopSensorPosM   := SEL(GVL_IHM.M1TreuilRetenue.Cmd.BtnHomingAtZero, _WinchM1CfgPersist.CfgTopSensorPos_M, 0.0),
    FwdRevSpeedFeedbackOff := HwIn.Winch.M1_ContactorsReleased_DI,
    BrakeFeedback        := HwIn.Winch.M1_BrakeIsOpen_DI,
    RawPos               := instEncoderAbsM1.RawPos,
    EncoderAvailable     := instEncoderAbsM1.EncoderAvailable,
    PresetAck            := instEncoderAbsM1.PresetAck,
    PresetNak            := instEncoderAbsM1.PresetNak,
    PointsPerRev         := 8192,
    MultiTurnRevsMax     := 4096,
    CableM_PerRev        := 2.0,
    BypassGlobal         := GVL_IHM.M1TreuilRetenue.Bypass.Global,
    Calib                := _CalibM1
);

instEncoderScaleM1(
    RawPos          := instEncoderAbsM1.RawPos,
    HomingRefRaw    := instHomingM1.HomingRefRaw,
    CableM_PerRev   := 2.0,
    PointsPerRev    := 8192
);

// 🧲 Codeurs M2 : Abs → Homing → Scale
instEncoderAbsM2(
    Enable              := TRUE,
    Reset               := PRG_SUPERVISION_CFC.FaultMachineReset_IHM,
    PowerContactorEngaged     := HwIn.Machine.PowerContactorEngaged_DI,
    Mode                := PRG_MODES_CFC.Auth.Mode,
    RawPosIn            := HwIn.Winch.COD2_PosValue,
    AlarmsIn            := HwIn.Winch.COD2_Alarms,
    WarningsIn          := HwIn.Winch.COD2_Warnings,
    SlaveOperational    := PRG_01_Diagnostics.instDiagEthercat.DeviceEncoderM2.Operational,
    PresetRequest       := instHomingM2.PresetRequest,
    PresetValue         := instHomingM2.PresetValue
);

instHomingM2(
    Enable               := TRUE,
    Reset                := PRG_SUPERVISION_CFC.FaultMachineReset_IHM,
    PowerContactorEngaged      := HwIn.Machine.PowerContactorEngaged_DI,
    Mode                 := PRG_MODES_CFC.Auth.Mode,
    Home                 := GVL_IHM.M2TreuilBenne.Cmd.BtnHome OR GVL_IHM.M2TreuilBenne.Cmd.BtnHomingAtZero,
    UnitaryMode          := (PRG_MODES_CFC.Auth.Mode = E_Mode.MAINT_N2)
                            AND (PRG_MODES_CFC.Auth.JoystickWinchSelectArbitrated <> 3),
    WinchSelected        := (PRG_MODES_CFC.Auth.JoystickWinchSelectArbitrated = 2),
    CfgHomingTargetM        := _WinchM2CfgPersist.CfgHomingTarget_M,
    BtnConfirmCoherence     := GVL_IHM.M2TreuilBenne.Cmd.BtnConfirmCoherence,
    TopPositionSensor    := HwIn.Winch.M1M2_TopPositionFree_DI,
    CfgTopSensorPosM   := SEL(GVL_IHM.M2TreuilBenne.Cmd.BtnHomingAtZero, _WinchM2CfgPersist.CfgTopSensorPos_M, 0.0),
    FwdRevSpeedFeedbackOff := HwIn.Winch.M2_ContactorsReleased_DI,
    BrakeFeedback        := HwIn.Winch.M2_BrakeIsOpen_DI,
    RawPos               := instEncoderAbsM2.RawPos,
    EncoderAvailable     := instEncoderAbsM2.EncoderAvailable,
    PresetAck            := instEncoderAbsM2.PresetAck,
    PresetNak            := instEncoderAbsM2.PresetNak,
    PointsPerRev         := 8192,
    MultiTurnRevsMax     := 4096,
    CableM_PerRev        := 2.0,
    BypassGlobal         := GVL_IHM.M2TreuilBenne.Bypass.Global,
    Calib                := _CalibM2
);

instEncoderScaleM2(
    RawPos          := instEncoderAbsM2.RawPos,
    HomingRefRaw    := instHomingM2.HomingRefRaw,
    CableM_PerRev   := 2.0,
    PointsPerRev    := 8192
);

// ↔️ Translation M3 : décodage du mot de capteurs de position
instPosDecoderM3(
    SensorTremie      := HwIn.Translation.M3_PosTremie_DI,
    SensorPV          := HwIn.Translation.M3_PosPV_DI,
    SensorP2          := HwIn.Translation.M3_PosP2_DI,
    SensorP1          := HwIn.Translation.M3_PosP1_DI,
    SensorMaintenance := HwIn.Translation.M3_PosMaintenance_DI
);

// 🆕 Exposition des positions Translation M3 pour les consommateurs legacy
TranslationPosTremie      := instPosDecoderM3.TranslationPosTremie;
TranslationPosPV          := instPosDecoderM3.TranslationPosPV;
TranslationPosP2          := instPosDecoderM3.TranslationPosP2;
TranslationPosP1          := instPosDecoderM3.TranslationPosP1;
TranslationPosMaintenance := instPosDecoderM3.TranslationPosMaintenance;

// 🆕 Filtrage PT1 (T#0MS = pass-through) des retours variateur M3 — cohérent avec le legacy
instCycleTimeAcq(DefaultValueS := 0.010);

instFilterM3StatusWord(
    ValueIn    := UINT_TO_REAL(WORD_TO_UINT(HwIn.Translation.M3_StatusWord)),
    TimeConst  := T#0MS,
    CycleTimeS := instCycleTimeAcq.CycleTimeS
);
M3_StatusWord_Filtered := REAL_TO_UINT(instFilterM3StatusWord.ValueOut);

instFilterM3ActualFreqHz(
    ValueIn    := UINT_TO_REAL(HwIn.Translation.M3_ActualFrequencyHz),
    TimeConst  := T#0MS,
    CycleTimeS := instCycleTimeAcq.CycleTimeS
);
M3_ActualFrequencyHz_Filtered := REAL_TO_UINT(instFilterM3ActualFreqHz.ValueOut);
